Fanuc KAREL source: kb00192.compact.KL

PROGRAM KB00192
%STACKSIZE=65535
%PRIORITY=65535
%NOLOCKGROUP
VAR
P1 : REAL
RESULT : INTEGER
BEGIN
P1=1.0
RESULT=TRUNC(P1)
END KB00192
